// #83: why F_CommandAcceptance rejected a command.
{attribute 'qualified_only'}
{attribute 'strict'}
TYPE E_CommandRejectReason :
(
	none := 0,
	estop,
	error,
	clock_invalid,
	stopping,
	powering_on,
	parking,
	parked,
	not_ready,
	gohome_active,
	init_required		// #72: manual mode since the last completed startup, send power=1 first
);
END_TYPE

(* stored: Version 1.1.0.1, ProductVersion 3.1.4024.15
   DUT E_CommandRejectReason: Id {5b1d2a10-7c3e-4d52-9a61-0e4f8c2b7a02} *)
